// TIA Portal V19 export
FUNCTION_BLOCK "RUA_R18"   // FB38, LAD
{ S7_Optimized_Access := 'TRUE' }
// stored: MemoryReserve 100, SetENOAutomatically false
   VAR
      START_Instance { S7_SetPoint := 'True'} : "START";
      "HEAT/COOL_Instance" { S7_SetPoint := 'True'} : "HEAT/COOL";
      "AUTO_COOLING_UTIITY SELECTION_Instance" { S7_SetPoint := 'True'} : "AUTO_COOLING_UTIITY SELECTION";
      AUTO_HEATING_SELECTION_Instance { S7_SetPoint := 'True'} : "AUTO_HEATING_SELECTION";
      COOLING_PROCESS_Instance { S7_SetPoint := 'True'} : "COOLING_PROCESS";
      "SEMI/_AUTO_Instance" { S7_SetPoint := 'True'} : "SEMI/_AUTO";
      HEATING_PROCEES_Instance { S7_SetPoint := 'True'} : "HEATING_PROCEES";
      RAMP_Instance { S7_SetPoint := 'True'} : "RAMP";
   END_VAR
BEGIN

REGION Network 1: START
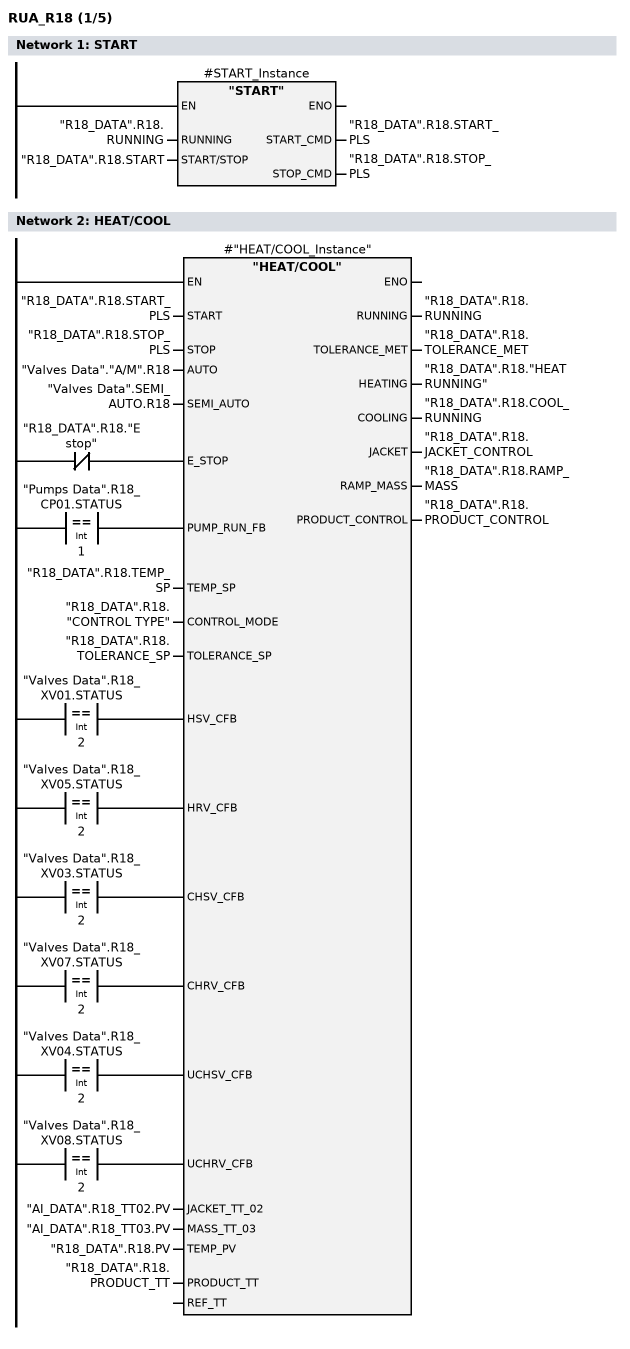
   RUNG wire#powerrail
      #START_Instance(RUNNING := "R18_DATA".R18.RUNNING, "START/STOP" := "R18_DATA".R18.START, START_CMD => "R18_DATA".R18.START_PLS, STOP_CMD => "R18_DATA".R18.STOP_PLS)
   END_RUNG
   // the same network as SCL:
   #START_Instance(RUNNING := "R18_DATA".R18.RUNNING,   // "START"
                   "START/STOP" := "R18_DATA".R18.START,
                   START_CMD => "R18_DATA".R18.START_PLS,
                   STOP_CMD => "R18_DATA".R18.STOP_PLS);
END_REGION

REGION Network 2: HEAT/COOL
   RUNG wire#powerrail
      #"HEAT/COOL_Instance"(E_STOP := wire#w1, PUMP_RUN_FB := wire#w2, HSV_CFB := wire#w3, HRV_CFB := wire#w4, CHSV_CFB := wire#w5, CHRV_CFB := wire#w6, UCHSV_CFB := wire#w7, UCHRV_CFB := wire#w8, START := "R18_DATA".R18.START_PLS, STOP := "R18_DATA".R18.STOP_PLS, AUTO := "Valves Data"."A/M".R18, SEMI_AUTO := "Valves Data".SEMI_AUTO.R18, TEMP_SP := "R18_DATA".R18.TEMP_SP, CONTROL_MODE := "R18_DATA".R18."CONTROL TYPE", TOLERANCE_SP := "R18_DATA".R18.TOLERANCE_SP, JACKET_TT_02 := "AI_DATA".R18_TT02.PV, MASS_TT_03 := "AI_DATA".R18_TT03.PV, TEMP_PV := "R18_DATA".R18.PV, PRODUCT_TT := "R18_DATA".R18.PRODUCT_TT, REF_TT :=, RUNNING => "R18_DATA".R18.RUNNING, TOLERANCE_MET => "R18_DATA".R18.TOLERANCE_MET, HEATING => "R18_DATA".R18."HEAT RUNNING", COOLING => "R18_DATA".R18.COOL_RUNNING, JACKET => "R18_DATA".R18.JACKET_CONTROL, RAMP_MASS => "R18_DATA".R18.RAMP_MASS, PRODUCT_CONTROL => "R18_DATA".R18.PRODUCT_CONTROL)
   END_RUNG
   RUNG wire#powerrail
      I_Contact( "R18_DATA".R18."E stop" )
   END_RUNG wire#w1
   RUNG wire#powerrail
      { S7_Templates := "SrcType := Int" } EQ_Contact(in1 := "Pumps Data".R18_CP01.STATUS, in2 := 1)
   END_RUNG wire#w2
   RUNG wire#powerrail
      { S7_Templates := "SrcType := Int" } EQ_Contact(in1 := "Valves Data".R18_XV01.STATUS, in2 := 2)
   END_RUNG wire#w3
   RUNG wire#powerrail
      { S7_Templates := "SrcType := Int" } EQ_Contact(in1 := "Valves Data".R18_XV05.STATUS, in2 := 2)
   END_RUNG wire#w4
   RUNG wire#powerrail
      { S7_Templates := "SrcType := Int" } EQ_Contact(in1 := "Valves Data".R18_XV03.STATUS, in2 := 2)
   END_RUNG wire#w5
   RUNG wire#powerrail
      { S7_Templates := "SrcType := Int" } EQ_Contact(in1 := "Valves Data".R18_XV07.STATUS, in2 := 2)
   END_RUNG wire#w6
   RUNG wire#powerrail
      { S7_Templates := "SrcType := Int" } EQ_Contact(in1 := "Valves Data".R18_XV04.STATUS, in2 := 2)
   END_RUNG wire#w7
   RUNG wire#powerrail
      { S7_Templates := "SrcType := Int" } EQ_Contact(in1 := "Valves Data".R18_XV08.STATUS, in2 := 2)
   END_RUNG wire#w8
   // the same network as SCL:
   #"HEAT/COOL_Instance"(START := "R18_DATA".R18.START_PLS,   // "HEAT/COOL"
                         STOP := "R18_DATA".R18.STOP_PLS,
                         AUTO := "Valves Data"."A/M".R18,
                         SEMI_AUTO := "Valves Data".SEMI_AUTO.R18,
                         E_STOP := NOT "R18_DATA".R18."E stop",
                         PUMP_RUN_FB := "Pumps Data".R18_CP01.STATUS = 1,
                         TEMP_SP := "R18_DATA".R18.TEMP_SP,
                         CONTROL_MODE := "R18_DATA".R18."CONTROL TYPE",
                         TOLERANCE_SP := "R18_DATA".R18.TOLERANCE_SP,
                         HSV_CFB := "Valves Data".R18_XV01.STATUS = 2,
                         HRV_CFB := "Valves Data".R18_XV05.STATUS = 2,
                         CHSV_CFB := "Valves Data".R18_XV03.STATUS = 2,
                         CHRV_CFB := "Valves Data".R18_XV07.STATUS = 2,
                         UCHSV_CFB := "Valves Data".R18_XV04.STATUS = 2,
                         UCHRV_CFB := "Valves Data".R18_XV08.STATUS = 2,
                         JACKET_TT_02 := "AI_DATA".R18_TT02.PV,
                         MASS_TT_03 := "AI_DATA".R18_TT03.PV,
                         TEMP_PV := "R18_DATA".R18.PV,
                         PRODUCT_TT := "R18_DATA".R18.PRODUCT_TT,
                         RUNNING => "R18_DATA".R18.RUNNING,
                         TOLERANCE_MET => "R18_DATA".R18.TOLERANCE_MET,
                         HEATING => "R18_DATA".R18."HEAT RUNNING",
                         COOLING => "R18_DATA".R18.COOL_RUNNING,
                         JACKET => "R18_DATA".R18.JACKET_CONTROL,
                         RAMP_MASS => "R18_DATA".R18.RAMP_MASS,
                         PRODUCT_CONTROL => "R18_DATA".R18.PRODUCT_CONTROL);
END_REGION

REGION Network 3: AUTO_COOLING
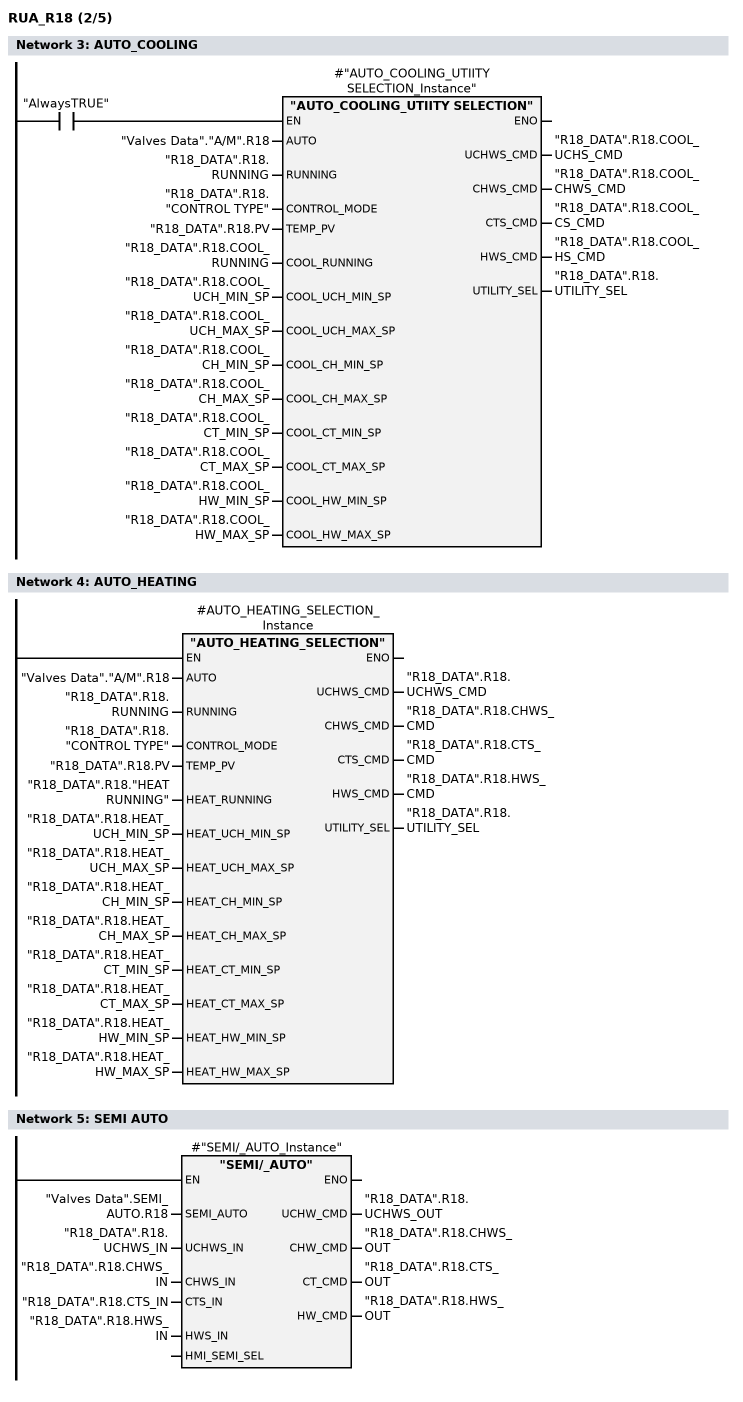
   RUNG wire#powerrail
      Contact( "AlwaysTRUE" )
      #"AUTO_COOLING_UTIITY SELECTION_Instance"(AUTO := "Valves Data"."A/M".R18, RUNNING := "R18_DATA".R18.RUNNING, CONTROL_MODE := "R18_DATA".R18."CONTROL TYPE", TEMP_PV := "R18_DATA".R18.PV, COOL_RUNNING := "R18_DATA".R18.COOL_RUNNING, COOL_UCH_MIN_SP := "R18_DATA".R18.COOL_UCH_MIN_SP, COOL_UCH_MAX_SP := "R18_DATA".R18.COOL_UCH_MAX_SP, COOL_CH_MIN_SP := "R18_DATA".R18.COOL_CH_MIN_SP, COOL_CH_MAX_SP := "R18_DATA".R18.COOL_CH_MAX_SP, COOL_CT_MIN_SP := "R18_DATA".R18.COOL_CT_MIN_SP, COOL_CT_MAX_SP := "R18_DATA".R18.COOL_CT_MAX_SP, COOL_HW_MIN_SP := "R18_DATA".R18.COOL_HW_MIN_SP, COOL_HW_MAX_SP := "R18_DATA".R18.COOL_HW_MAX_SP, UCHWS_CMD => "R18_DATA".R18.COOL_UCHS_CMD, CHWS_CMD => "R18_DATA".R18.COOL_CHWS_CMD, CTS_CMD => "R18_DATA".R18.COOL_CS_CMD, HWS_CMD => "R18_DATA".R18.COOL_HS_CMD, UTILITY_SEL => "R18_DATA".R18.UTILITY_SEL)
   END_RUNG
   // the same network as SCL:
   IF "AlwaysTRUE" THEN
       #"AUTO_COOLING_UTIITY SELECTION_Instance"(AUTO := "Valves Data"."A/M".R18,   // "AUTO_COOLING_UTIITY SELECTION"
                               RUNNING := "R18_DATA".R18.RUNNING,
                               CONTROL_MODE := "R18_DATA".R18."CONTROL TYPE",
                               TEMP_PV := "R18_DATA".R18.PV,
                               COOL_RUNNING := "R18_DATA".R18.COOL_RUNNING,
                               COOL_UCH_MIN_SP := "R18_DATA".R18.COOL_UCH_MIN_SP,
                               COOL_UCH_MAX_SP := "R18_DATA".R18.COOL_UCH_MAX_SP,
                               COOL_CH_MIN_SP := "R18_DATA".R18.COOL_CH_MIN_SP,
                               COOL_CH_MAX_SP := "R18_DATA".R18.COOL_CH_MAX_SP,
                               COOL_CT_MIN_SP := "R18_DATA".R18.COOL_CT_MIN_SP,
                               COOL_CT_MAX_SP := "R18_DATA".R18.COOL_CT_MAX_SP,
                               COOL_HW_MIN_SP := "R18_DATA".R18.COOL_HW_MIN_SP,
                               COOL_HW_MAX_SP := "R18_DATA".R18.COOL_HW_MAX_SP,
                               UCHWS_CMD => "R18_DATA".R18.COOL_UCHS_CMD,
                               CHWS_CMD => "R18_DATA".R18.COOL_CHWS_CMD,
                               CTS_CMD => "R18_DATA".R18.COOL_CS_CMD,
                               HWS_CMD => "R18_DATA".R18.COOL_HS_CMD,
                               UTILITY_SEL => "R18_DATA".R18.UTILITY_SEL);
   END_IF;
END_REGION

REGION Network 4: AUTO_HEATING
   RUNG wire#powerrail
      #AUTO_HEATING_SELECTION_Instance(AUTO := "Valves Data"."A/M".R18, RUNNING := "R18_DATA".R18.RUNNING, CONTROL_MODE := "R18_DATA".R18."CONTROL TYPE", TEMP_PV := "R18_DATA".R18.PV, HEAT_RUNNING := "R18_DATA".R18."HEAT RUNNING", HEAT_UCH_MIN_SP := "R18_DATA".R18.HEAT_UCH_MIN_SP, HEAT_UCH_MAX_SP := "R18_DATA".R18.HEAT_UCH_MAX_SP, HEAT_CH_MIN_SP := "R18_DATA".R18.HEAT_CH_MIN_SP, HEAT_CH_MAX_SP := "R18_DATA".R18.HEAT_CH_MAX_SP, HEAT_CT_MIN_SP := "R18_DATA".R18.HEAT_CT_MIN_SP, HEAT_CT_MAX_SP := "R18_DATA".R18.HEAT_CT_MAX_SP, HEAT_HW_MIN_SP := "R18_DATA".R18.HEAT_HW_MIN_SP, HEAT_HW_MAX_SP := "R18_DATA".R18.HEAT_HW_MAX_SP, UCHWS_CMD => "R18_DATA".R18.UCHWS_CMD, CHWS_CMD => "R18_DATA".R18.CHWS_CMD, CTS_CMD => "R18_DATA".R18.CTS_CMD, HWS_CMD => "R18_DATA".R18.HWS_CMD, UTILITY_SEL => "R18_DATA".R18.UTILITY_SEL)
   END_RUNG
   // the same network as SCL:
   #AUTO_HEATING_SELECTION_Instance(AUTO := "Valves Data"."A/M".R18,   // "AUTO_HEATING_SELECTION"
                           RUNNING := "R18_DATA".R18.RUNNING,
                           CONTROL_MODE := "R18_DATA".R18."CONTROL TYPE",
                           TEMP_PV := "R18_DATA".R18.PV,
                           HEAT_RUNNING := "R18_DATA".R18."HEAT RUNNING",
                           HEAT_UCH_MIN_SP := "R18_DATA".R18.HEAT_UCH_MIN_SP,
                           HEAT_UCH_MAX_SP := "R18_DATA".R18.HEAT_UCH_MAX_SP,
                           HEAT_CH_MIN_SP := "R18_DATA".R18.HEAT_CH_MIN_SP,
                           HEAT_CH_MAX_SP := "R18_DATA".R18.HEAT_CH_MAX_SP,
                           HEAT_CT_MIN_SP := "R18_DATA".R18.HEAT_CT_MIN_SP,
                           HEAT_CT_MAX_SP := "R18_DATA".R18.HEAT_CT_MAX_SP,
                           HEAT_HW_MIN_SP := "R18_DATA".R18.HEAT_HW_MIN_SP,
                           HEAT_HW_MAX_SP := "R18_DATA".R18.HEAT_HW_MAX_SP,
                           UCHWS_CMD => "R18_DATA".R18.UCHWS_CMD,
                           CHWS_CMD => "R18_DATA".R18.CHWS_CMD,
                           CTS_CMD => "R18_DATA".R18.CTS_CMD,
                           HWS_CMD => "R18_DATA".R18.HWS_CMD,
                           UTILITY_SEL => "R18_DATA".R18.UTILITY_SEL);
END_REGION

REGION Network 5: SEMI AUTO
   RUNG wire#powerrail
      #"SEMI/_AUTO_Instance"(SEMI_AUTO := "Valves Data".SEMI_AUTO.R18, UCHWS_IN := "R18_DATA".R18.UCHWS_IN, CHWS_IN := "R18_DATA".R18.CHWS_IN, CTS_IN := "R18_DATA".R18.CTS_IN, HWS_IN := "R18_DATA".R18.HWS_IN, UCHW_CMD => "R18_DATA".R18.UCHWS_OUT, CHW_CMD => "R18_DATA".R18.CHWS_OUT, CT_CMD => "R18_DATA".R18.CTS_OUT, HW_CMD => "R18_DATA".R18.HWS_OUT, HMI_SEMI_SEL :=)
   END_RUNG
   // the same network as SCL:
   #"SEMI/_AUTO_Instance"(SEMI_AUTO := "Valves Data".SEMI_AUTO.R18,   // "SEMI/_AUTO"
                          UCHWS_IN := "R18_DATA".R18.UCHWS_IN,
                          CHWS_IN := "R18_DATA".R18.CHWS_IN,
                          CTS_IN := "R18_DATA".R18.CTS_IN,
                          HWS_IN := "R18_DATA".R18.HWS_IN,
                          UCHW_CMD => "R18_DATA".R18.UCHWS_OUT,
                          CHW_CMD => "R18_DATA".R18.CHWS_OUT,
                          CT_CMD => "R18_DATA".R18.CTS_OUT,
                          HW_CMD => "R18_DATA".R18.HWS_OUT);
END_REGION

REGION Network 6: COOLING_PROCESS
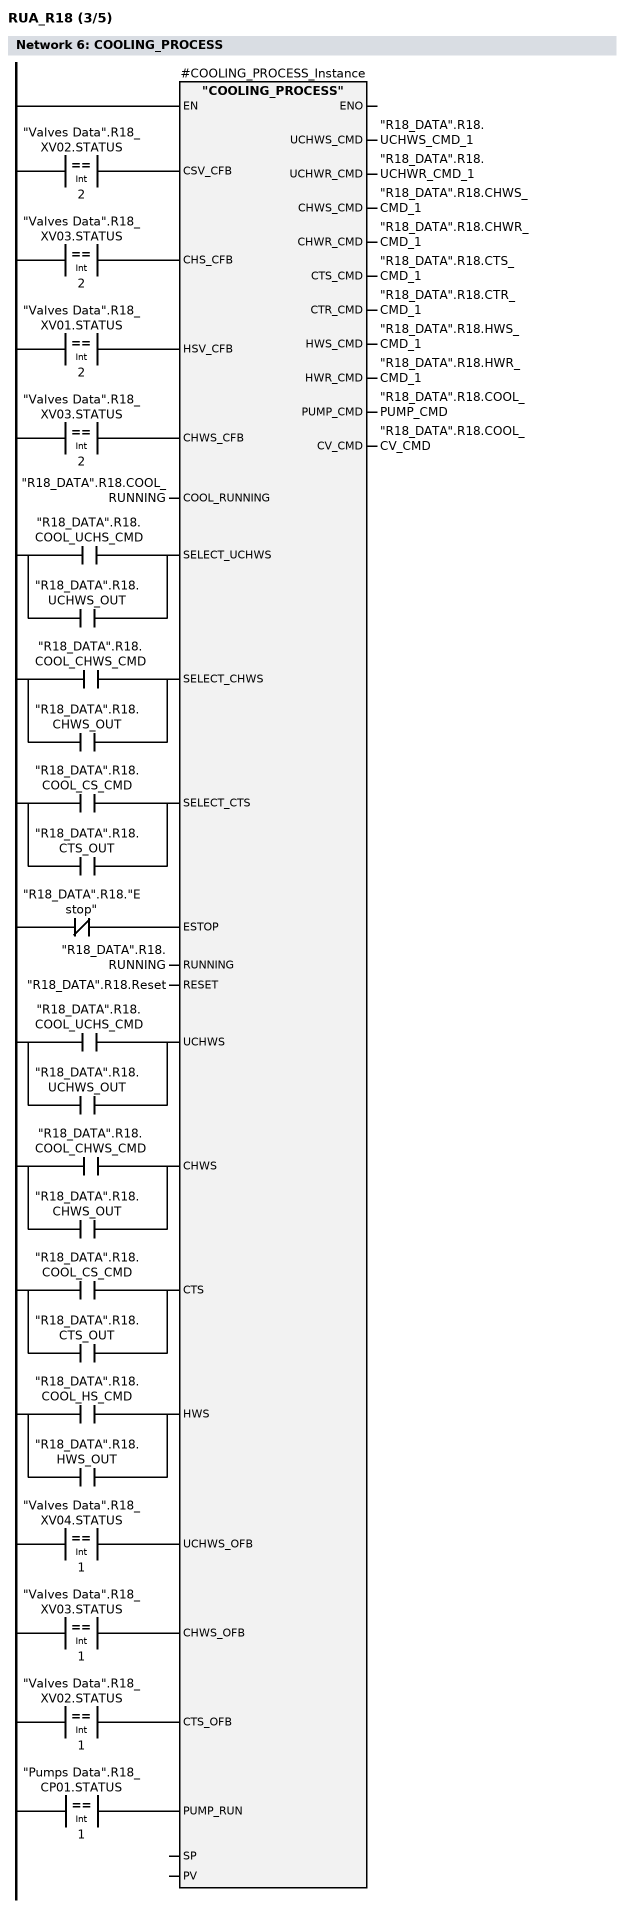
   RUNG wire#powerrail
      #COOLING_PROCESS_Instance(CSV_CFB := wire#w1, CHS_CFB := wire#w2, HSV_CFB := wire#w3, CHWS_CFB := wire#w4, SELECT_UCHWS := wire#w5, SELECT_CHWS := wire#w6, SELECT_CTS := wire#w7, ESTOP := wire#w8, UCHWS := wire#w9, CHWS := wire#w10, CTS := wire#w11, HWS := wire#w12, UCHWS_OFB := wire#w13, CHWS_OFB := wire#w14, CTS_OFB := wire#w15, PUMP_RUN := wire#w16, COOL_RUNNING := "R18_DATA".R18.COOL_RUNNING, RUNNING := "R18_DATA".R18.RUNNING, RESET := "R18_DATA".R18.Reset, SP :=, PV :=, UCHWS_CMD => "R18_DATA".R18.UCHWS_CMD_1, UCHWR_CMD => "R18_DATA".R18.UCHWR_CMD_1, CHWS_CMD => "R18_DATA".R18.CHWS_CMD_1, CHWR_CMD => "R18_DATA".R18.CHWR_CMD_1, CTS_CMD => "R18_DATA".R18.CTS_CMD_1, CTR_CMD => "R18_DATA".R18.CTR_CMD_1, HWS_CMD => "R18_DATA".R18.HWS_CMD_1, HWR_CMD => "R18_DATA".R18.HWR_CMD_1, PUMP_CMD => "R18_DATA".R18.COOL_PUMP_CMD, CV_CMD => "R18_DATA".R18.COOL_CV_CMD)
   END_RUNG
   RUNG wire#powerrail
      { S7_Templates := "SrcType := Int" } EQ_Contact(in1 := "Valves Data".R18_XV02.STATUS, in2 := 2)
   END_RUNG wire#w1
   RUNG wire#powerrail
      { S7_Templates := "SrcType := Int" } EQ_Contact(in1 := "Valves Data".R18_XV03.STATUS, in2 := 2)
   END_RUNG wire#w2
   RUNG wire#powerrail
      { S7_Templates := "SrcType := Int" } EQ_Contact(in1 := "Valves Data".R18_XV01.STATUS, in2 := 2)
   END_RUNG wire#w3
   RUNG wire#powerrail
      { S7_Templates := "SrcType := Int" } EQ_Contact(in1 := "Valves Data".R18_XV03.STATUS, in2 := 2)
   END_RUNG wire#w4
   RUNG wire#powerrail
      Contact( "R18_DATA".R18.COOL_UCHS_CMD )
   END_RUNG wire#w5
   RUNG wire#powerrail
      Contact( "R18_DATA".R18.UCHWS_OUT )
   END_RUNG wire#w5
   RUNG wire#powerrail
      Contact( "R18_DATA".R18.COOL_CHWS_CMD )
   END_RUNG wire#w6
   RUNG wire#powerrail
      Contact( "R18_DATA".R18.CHWS_OUT )
   END_RUNG wire#w6
   RUNG wire#powerrail
      Contact( "R18_DATA".R18.COOL_CS_CMD )
   END_RUNG wire#w7
   RUNG wire#powerrail
      Contact( "R18_DATA".R18.CTS_OUT )
   END_RUNG wire#w7
   RUNG wire#powerrail
      I_Contact( "R18_DATA".R18."E stop" )
   END_RUNG wire#w8
   RUNG wire#powerrail
      Contact( "R18_DATA".R18.COOL_UCHS_CMD )
   END_RUNG wire#w9
   RUNG wire#powerrail
      Contact( "R18_DATA".R18.UCHWS_OUT )
   END_RUNG wire#w9
   RUNG wire#powerrail
      Contact( "R18_DATA".R18.COOL_CHWS_CMD )
   END_RUNG wire#w10
   RUNG wire#powerrail
      Contact( "R18_DATA".R18.CHWS_OUT )
   END_RUNG wire#w10
   RUNG wire#powerrail
      Contact( "R18_DATA".R18.COOL_CS_CMD )
   END_RUNG wire#w11
   RUNG wire#powerrail
      Contact( "R18_DATA".R18.CTS_OUT )
   END_RUNG wire#w11
   RUNG wire#powerrail
      Contact( "R18_DATA".R18.COOL_HS_CMD )
   END_RUNG wire#w12
   RUNG wire#powerrail
      Contact( "R18_DATA".R18.HWS_OUT )
   END_RUNG wire#w12
   RUNG wire#powerrail
      { S7_Templates := "SrcType := Int" } EQ_Contact(in1 := "Valves Data".R18_XV04.STATUS, in2 := 1)
   END_RUNG wire#w13
   RUNG wire#powerrail
      { S7_Templates := "SrcType := Int" } EQ_Contact(in1 := "Valves Data".R18_XV03.STATUS, in2 := 1)
   END_RUNG wire#w14
   RUNG wire#powerrail
      { S7_Templates := "SrcType := Int" } EQ_Contact(in1 := "Valves Data".R18_XV02.STATUS, in2 := 1)
   END_RUNG wire#w15
   RUNG wire#powerrail
      { S7_Templates := "SrcType := Int" } EQ_Contact(in1 := "Pumps Data".R18_CP01.STATUS, in2 := 1)
   END_RUNG wire#w16
   // the same network as SCL:
   #COOLING_PROCESS_Instance(CSV_CFB := "Valves Data".R18_XV02.STATUS = 2,   // "COOLING_PROCESS"
                           CHS_CFB := "Valves Data".R18_XV03.STATUS = 2,
                           HSV_CFB := "Valves Data".R18_XV01.STATUS = 2,
                           CHWS_CFB := "Valves Data".R18_XV03.STATUS = 2,
                           COOL_RUNNING := "R18_DATA".R18.COOL_RUNNING,
                           SELECT_UCHWS := "R18_DATA".R18.COOL_UCHS_CMD OR "R18_DATA".R18.UCHWS_OUT,
                           SELECT_CHWS := "R18_DATA".R18.COOL_CHWS_CMD OR "R18_DATA".R18.CHWS_OUT,
                           SELECT_CTS := "R18_DATA".R18.COOL_CS_CMD OR "R18_DATA".R18.CTS_OUT,
                           ESTOP := NOT "R18_DATA".R18."E stop",
                           RUNNING := "R18_DATA".R18.RUNNING,
                           RESET := "R18_DATA".R18.Reset,
                           UCHWS := "R18_DATA".R18.COOL_UCHS_CMD OR "R18_DATA".R18.UCHWS_OUT,
                           CHWS := "R18_DATA".R18.COOL_CHWS_CMD OR "R18_DATA".R18.CHWS_OUT,
                           CTS := "R18_DATA".R18.COOL_CS_CMD OR "R18_DATA".R18.CTS_OUT,
                           HWS := "R18_DATA".R18.COOL_HS_CMD OR "R18_DATA".R18.HWS_OUT,
                           UCHWS_OFB := "Valves Data".R18_XV04.STATUS = 1,
                           CHWS_OFB := "Valves Data".R18_XV03.STATUS = 1,
                           CTS_OFB := "Valves Data".R18_XV02.STATUS = 1,
                           PUMP_RUN := "Pumps Data".R18_CP01.STATUS = 1,
                           UCHWS_CMD => "R18_DATA".R18.UCHWS_CMD_1,
                           UCHWR_CMD => "R18_DATA".R18.UCHWR_CMD_1,
                           CHWS_CMD => "R18_DATA".R18.CHWS_CMD_1,
                           CHWR_CMD => "R18_DATA".R18.CHWR_CMD_1,
                           CTS_CMD => "R18_DATA".R18.CTS_CMD_1,
                           CTR_CMD => "R18_DATA".R18.CTR_CMD_1,
                           HWS_CMD => "R18_DATA".R18.HWS_CMD_1,
                           HWR_CMD => "R18_DATA".R18.HWR_CMD_1,
                           PUMP_CMD => "R18_DATA".R18.COOL_PUMP_CMD,
                           CV_CMD => "R18_DATA".R18.COOL_CV_CMD);
END_REGION

REGION Network 7: HEATING PROCESS
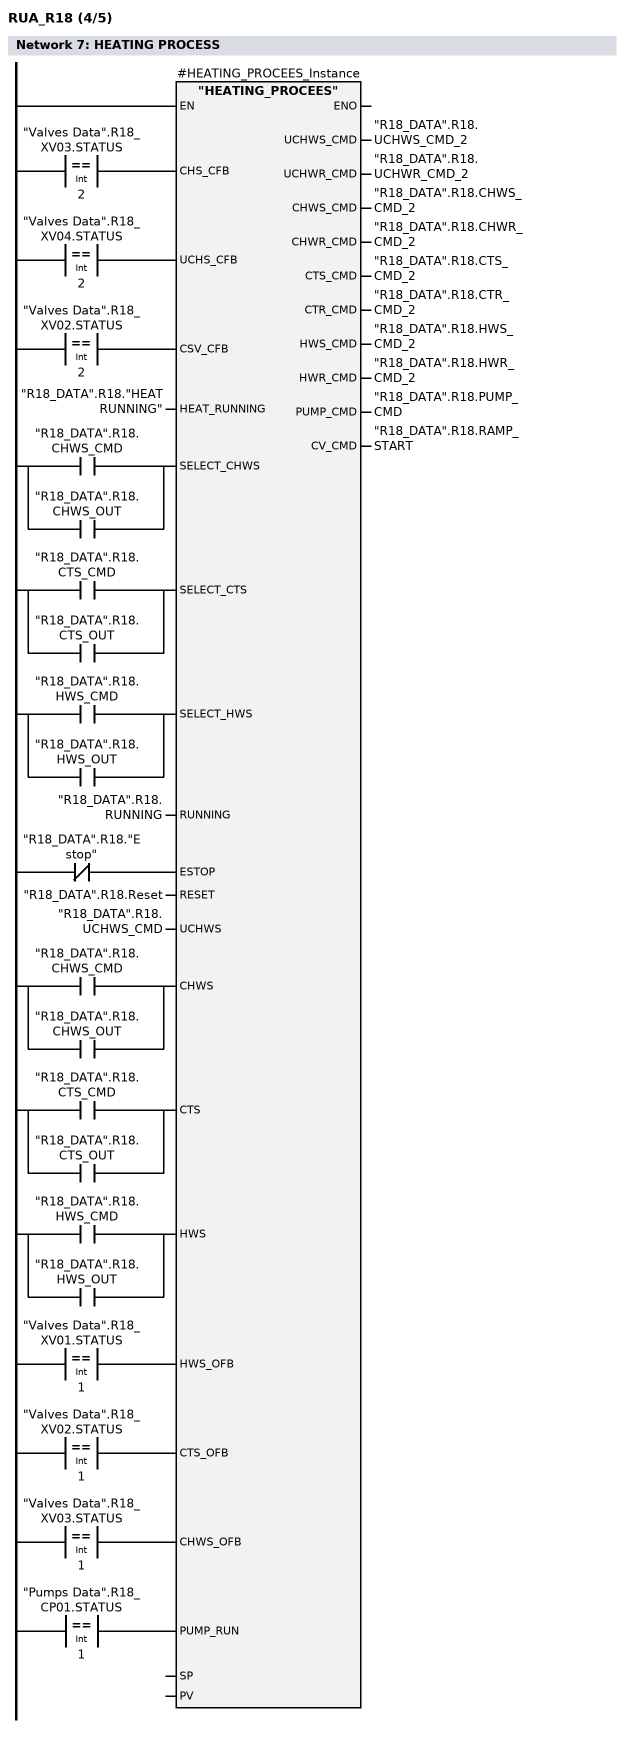
   RUNG wire#powerrail
      #HEATING_PROCEES_Instance(CHS_CFB := wire#w1, UCHS_CFB := wire#w2, CSV_CFB := wire#w3, SELECT_CHWS := wire#w4, SELECT_CTS := wire#w5, SELECT_HWS := wire#w6, ESTOP := wire#w7, CHWS := wire#w8, CTS := wire#w9, HWS := wire#w10, HWS_OFB := wire#w11, CTS_OFB := wire#w12, CHWS_OFB := wire#w13, PUMP_RUN := wire#w14, HEAT_RUNNING := "R18_DATA".R18."HEAT RUNNING", RUNNING := "R18_DATA".R18.RUNNING, RESET := "R18_DATA".R18.Reset, UCHWS := "R18_DATA".R18.UCHWS_CMD, SP :=, PV :=, UCHWS_CMD => "R18_DATA".R18.UCHWS_CMD_2, UCHWR_CMD => "R18_DATA".R18.UCHWR_CMD_2, CHWS_CMD => "R18_DATA".R18.CHWS_CMD_2, CHWR_CMD => "R18_DATA".R18.CHWR_CMD_2, CTS_CMD => "R18_DATA".R18.CTS_CMD_2, CTR_CMD => "R18_DATA".R18.CTR_CMD_2, HWS_CMD => "R18_DATA".R18.HWS_CMD_2, HWR_CMD => "R18_DATA".R18.HWR_CMD_2, PUMP_CMD => "R18_DATA".R18.PUMP_CMD, CV_CMD => "R18_DATA".R18.RAMP_START)
   END_RUNG
   RUNG wire#powerrail
      { S7_Templates := "SrcType := Int" } EQ_Contact(in1 := "Valves Data".R18_XV03.STATUS, in2 := 2)
   END_RUNG wire#w1
   RUNG wire#powerrail
      { S7_Templates := "SrcType := Int" } EQ_Contact(in1 := "Valves Data".R18_XV04.STATUS, in2 := 2)
   END_RUNG wire#w2
   RUNG wire#powerrail
      { S7_Templates := "SrcType := Int" } EQ_Contact(in1 := "Valves Data".R18_XV02.STATUS, in2 := 2)
   END_RUNG wire#w3
   RUNG wire#powerrail
      Contact( "R18_DATA".R18.CHWS_CMD )
   END_RUNG wire#w4
   RUNG wire#powerrail
      Contact( "R18_DATA".R18.CHWS_OUT )
   END_RUNG wire#w4
   RUNG wire#powerrail
      Contact( "R18_DATA".R18.CTS_CMD )
   END_RUNG wire#w5
   RUNG wire#powerrail
      Contact( "R18_DATA".R18.CTS_OUT )
   END_RUNG wire#w5
   RUNG wire#powerrail
      Contact( "R18_DATA".R18.HWS_CMD )
   END_RUNG wire#w6
   RUNG wire#powerrail
      Contact( "R18_DATA".R18.HWS_OUT )
   END_RUNG wire#w6
   RUNG wire#powerrail
      I_Contact( "R18_DATA".R18."E stop" )
   END_RUNG wire#w7
   RUNG wire#powerrail
      Contact( "R18_DATA".R18.CHWS_CMD )
   END_RUNG wire#w8
   RUNG wire#powerrail
      Contact( "R18_DATA".R18.CHWS_OUT )
   END_RUNG wire#w8
   RUNG wire#powerrail
      Contact( "R18_DATA".R18.CTS_CMD )
   END_RUNG wire#w9
   RUNG wire#powerrail
      Contact( "R18_DATA".R18.CTS_OUT )
   END_RUNG wire#w9
   RUNG wire#powerrail
      Contact( "R18_DATA".R18.HWS_CMD )
   END_RUNG wire#w10
   RUNG wire#powerrail
      Contact( "R18_DATA".R18.HWS_OUT )
   END_RUNG wire#w10
   RUNG wire#powerrail
      { S7_Templates := "SrcType := Int" } EQ_Contact(in1 := "Valves Data".R18_XV01.STATUS, in2 := 1)
   END_RUNG wire#w11
   RUNG wire#powerrail
      { S7_Templates := "SrcType := Int" } EQ_Contact(in1 := "Valves Data".R18_XV02.STATUS, in2 := 1)
   END_RUNG wire#w12
   RUNG wire#powerrail
      { S7_Templates := "SrcType := Int" } EQ_Contact(in1 := "Valves Data".R18_XV03.STATUS, in2 := 1)
   END_RUNG wire#w13
   RUNG wire#powerrail
      { S7_Templates := "SrcType := Int" } EQ_Contact(in1 := "Pumps Data".R18_CP01.STATUS, in2 := 1)
   END_RUNG wire#w14
   // the same network as SCL:
   #HEATING_PROCEES_Instance(CHS_CFB := "Valves Data".R18_XV03.STATUS = 2,   // "HEATING_PROCEES"
                           UCHS_CFB := "Valves Data".R18_XV04.STATUS = 2,
                           CSV_CFB := "Valves Data".R18_XV02.STATUS = 2,
                           HEAT_RUNNING := "R18_DATA".R18."HEAT RUNNING",
                           SELECT_CHWS := "R18_DATA".R18.CHWS_CMD OR "R18_DATA".R18.CHWS_OUT,
                           SELECT_CTS := "R18_DATA".R18.CTS_CMD OR "R18_DATA".R18.CTS_OUT,
                           SELECT_HWS := "R18_DATA".R18.HWS_CMD OR "R18_DATA".R18.HWS_OUT,
                           RUNNING := "R18_DATA".R18.RUNNING,
                           ESTOP := NOT "R18_DATA".R18."E stop",
                           RESET := "R18_DATA".R18.Reset,
                           UCHWS := "R18_DATA".R18.UCHWS_CMD,
                           CHWS := "R18_DATA".R18.CHWS_CMD OR "R18_DATA".R18.CHWS_OUT,
                           CTS := "R18_DATA".R18.CTS_CMD OR "R18_DATA".R18.CTS_OUT,
                           HWS := "R18_DATA".R18.HWS_CMD OR "R18_DATA".R18.HWS_OUT,
                           HWS_OFB := "Valves Data".R18_XV01.STATUS = 1,
                           CTS_OFB := "Valves Data".R18_XV02.STATUS = 1,
                           CHWS_OFB := "Valves Data".R18_XV03.STATUS = 1,
                           PUMP_RUN := "Pumps Data".R18_CP01.STATUS = 1,
                           UCHWS_CMD => "R18_DATA".R18.UCHWS_CMD_2,
                           UCHWR_CMD => "R18_DATA".R18.UCHWR_CMD_2,
                           CHWS_CMD => "R18_DATA".R18.CHWS_CMD_2,
                           CHWR_CMD => "R18_DATA".R18.CHWR_CMD_2,
                           CTS_CMD => "R18_DATA".R18.CTS_CMD_2,
                           CTR_CMD => "R18_DATA".R18.CTR_CMD_2,
                           HWS_CMD => "R18_DATA".R18.HWS_CMD_2,
                           HWR_CMD => "R18_DATA".R18.HWR_CMD_2,
                           PUMP_CMD => "R18_DATA".R18.PUMP_CMD,
                           CV_CMD => "R18_DATA".R18.RAMP_START);
END_REGION

REGION Network 8: RAMP
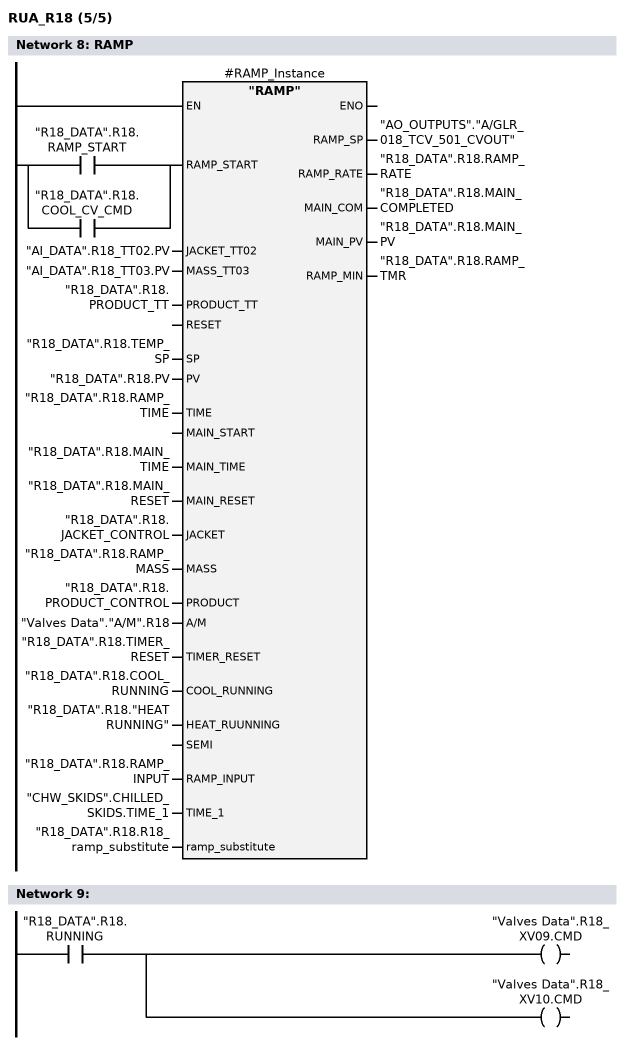
   RUNG wire#powerrail
      #RAMP_Instance(RAMP_START := wire#w1, JACKET_TT02 := "AI_DATA".R18_TT02.PV, MASS_TT03 := "AI_DATA".R18_TT03.PV, PRODUCT_TT := "R18_DATA".R18.PRODUCT_TT, RESET :=, SP := "R18_DATA".R18.TEMP_SP, PV := "R18_DATA".R18.PV, "TIME" := "R18_DATA".R18.RAMP_TIME, MAIN_START :=, MAIN_TIME := "R18_DATA".R18.MAIN_TIME, MAIN_RESET := "R18_DATA".R18.MAIN_RESET, JACKET := "R18_DATA".R18.JACKET_CONTROL, MASS := "R18_DATA".R18.RAMP_MASS, PRODUCT := "R18_DATA".R18.PRODUCT_CONTROL, "A/M" := "Valves Data"."A/M".R18, TIMER_RESET := "R18_DATA".R18.TIMER_RESET, COOL_RUNNING := "R18_DATA".R18.COOL_RUNNING, HEAT_RUUNNING := "R18_DATA".R18."HEAT RUNNING", RAMP_INPUT := "R18_DATA".R18.RAMP_INPUT, TIME_1 := "CHW_SKIDS".CHILLED_SKIDS.TIME_1, ramp_substitute := "R18_DATA".R18.R18_ramp_substitute, RAMP_SP => "AO_OUTPUTS"."A/GLR_018_TCV_501_CVOUT", RAMP_RATE => "R18_DATA".R18.RAMP_RATE, MAIN_COM => "R18_DATA".R18.MAIN_COMPLETED, MAIN_PV => "R18_DATA".R18.MAIN_PV, RAMP_MIN => "R18_DATA".R18.RAMP_TMR, SEMI :=)
   END_RUNG
   RUNG wire#powerrail
      Contact( "R18_DATA".R18.RAMP_START )
   END_RUNG wire#w1
   RUNG wire#powerrail
      Contact( "R18_DATA".R18.COOL_CV_CMD )
   END_RUNG wire#w1
   // the same network as SCL:
   #RAMP_Instance(RAMP_START := "R18_DATA".R18.RAMP_START OR "R18_DATA".R18.COOL_CV_CMD,   // "RAMP"
                  JACKET_TT02 := "AI_DATA".R18_TT02.PV,
                  MASS_TT03 := "AI_DATA".R18_TT03.PV,
                  PRODUCT_TT := "R18_DATA".R18.PRODUCT_TT,
                  SP := "R18_DATA".R18.TEMP_SP,
                  PV := "R18_DATA".R18.PV,
                  "TIME" := "R18_DATA".R18.RAMP_TIME,
                  MAIN_TIME := "R18_DATA".R18.MAIN_TIME,
                  MAIN_RESET := "R18_DATA".R18.MAIN_RESET,
                  JACKET := "R18_DATA".R18.JACKET_CONTROL,
                  MASS := "R18_DATA".R18.RAMP_MASS,
                  PRODUCT := "R18_DATA".R18.PRODUCT_CONTROL,
                  "A/M" := "Valves Data"."A/M".R18,
                  TIMER_RESET := "R18_DATA".R18.TIMER_RESET,
                  COOL_RUNNING := "R18_DATA".R18.COOL_RUNNING,
                  HEAT_RUUNNING := "R18_DATA".R18."HEAT RUNNING",
                  RAMP_INPUT := "R18_DATA".R18.RAMP_INPUT,
                  TIME_1 := "CHW_SKIDS".CHILLED_SKIDS.TIME_1,
                  ramp_substitute := "R18_DATA".R18.R18_ramp_substitute,
                  RAMP_SP => "AO_OUTPUTS"."A/GLR_018_TCV_501_CVOUT",
                  RAMP_RATE => "R18_DATA".R18.RAMP_RATE,
                  MAIN_COM => "R18_DATA".R18.MAIN_COMPLETED,
                  MAIN_PV => "R18_DATA".R18.MAIN_PV,
                  RAMP_MIN => "R18_DATA".R18.RAMP_TMR);
END_REGION

REGION Network 9
   RUNG wire#powerrail
      Contact( "R18_DATA".R18.RUNNING )
      wire#w1
      Coil( "Valves Data".R18_XV09.CMD )
   END_RUNG
   RUNG wire#w1
      Coil( "Valves Data".R18_XV10.CMD )
   END_RUNG
   // the same network as SCL:
   "Valves Data".R18_XV09.CMD := "R18_DATA".R18.RUNNING;
   "Valves Data".R18_XV10.CMD := "R18_DATA".R18.RUNNING;
END_REGION
END_FUNCTION_BLOCK
